(* IEC 61131-3 sources: IRIS-Project/LASAL CONTROL SOFTWARE/LasalProject_2025_09_12/Class/Rack12V, 1 file *)

(* ---- Rack12V.st ---- *)
(*!
<Class
	Name               = "Rack12V"
	Revision           = "0.0"
	RealtimeTask       = "false"
	CyclicTask         = "false"
	BackgroundTask     = "true"
	DefBackground      = "100 ms"
	Sigmatek           = "false"
	OSInterface        = "false"
	HighPriority       = "false"
	Automatic          = "false"
	UpdateMode         = "Prescan"
	SharedCommandTable = "true"
	Objectsize         = "(330,120)">
	<Channels>
		<Server Name="ClassSvr" Visualized="false" Initialize="false" WriteProtected="true" Retentive="false"/>
		<Server Name="Command_Rack" Visualized="false" Initialize="false" WriteProtected="false" Retentive="false"/>
		<Client Name="ToPLC" Required="true" Internal="false"/>
	</Channels>
</Class>
*)
Rack12V : CLASS
	TYPE
	  t_CommandRack :  //! <Type Public="true" Name="t_CommandRack"/>
	  (
	    Idle:=10,
	    Command_On:=1,
	    Command_Off:=0
	  )$UDINT;
	END_TYPE
  //Servers:
	ClassSvr 	: SvrChCmd_DINT;
	Command_Rack 	: SvrCh_t_CommandRack_PTofCls_Rack12V;
  //Clients:
	ToPLC 	: CltCh_DINT;
  //Variables:
		v_CaseRack12V 	: t_CommandRack;
  //Functions:

	FUNCTION VIRTUAL GLOBAL Init;

	FUNCTION VIRTUAL GLOBAL Background
		VAR_INPUT
			EAX 	: UDINT;
		END_VAR
		VAR_OUTPUT
			state (EAX) 	: UDINT;
		END_VAR;

	FUNCTION VIRTUAL GLOBAL Command_Rack::Read
		VAR_OUTPUT
			output (EAX) 	: Rack12V::t_CommandRack;
		END_VAR;
  //Tables:
	FUNCTION @STD
		VAR_OUTPUT
			ret_code	: CONFSTATES;
		END_VAR;
	FUNCTION GLOBAL TAB @CT_;
END_CLASS;

FUNCTION VIRTUAL GLOBAL Rack12V::Background
	VAR_INPUT
		EAX 	: UDINT;
	END_VAR
	VAR_OUTPUT
		state (EAX) 	: UDINT;
	END_VAR

  v_CaseRack12V:=Command_Rack.Read();

  case v_CaseRack12V of

    Idle:

    Command_Off:
      ToPLC.Write(input:=1);
      Command_Rack.Write(input:=Idle);

    Command_On:
      ToPLC.Write(input:=0);
      Command_Rack.Write(input:=Idle);

  end_case;

	state := READY;

END_FUNCTION

FUNCTION VIRTUAL GLOBAL Rack12V::Init
v_CaseRack12V:=Idle;

END_FUNCTION

FUNCTION VIRTUAL GLOBAL Rack12V::Command_Rack::Read
	VAR_OUTPUT
		output (EAX) 	: Rack12V::t_CommandRack;
	END_VAR

	output := Command_Rack;

END_FUNCTION
